SUBAPPLICATION GreenWhiteBackground2_AXC (* Hintergrundfarbe (TRUE -> Grün, FALSE -> Weiß) für 2 Objekte (AX-Adapter) (Kompakt) *)
  (* Standard: 61499-2 *)
  (* Version 1.0, 2026-07-21, franz, Meisterschulen am Ostbahnhof *)
  PACKAGE MyLib::sys;
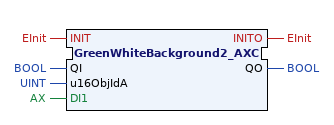
  EVENT_INPUT
    INIT : EInit; (* Initialization Request *)
  END_EVENT
  EVENT_OUTPUT
    INITO : EInit; (* Initialization Confirm *)
  END_EVENT
  VAR_INPUT
    QI : BOOL := TRUE; (* Quality Input - TRUE to enable service *)
    u16ObjIdA : UINT;
  END_VAR
  VAR_OUTPUT
    QO : BOOL; (* Quality Output - TRUE if service executed successfully *)
  END_VAR
  SOCKETS
    DI1 : adapter::types::unidirectional::AX;
  END_SOCKETS
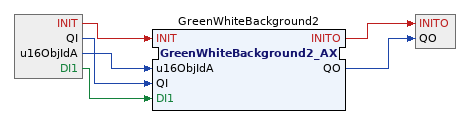
  SUBAPPS
    GreenWhiteBackground2 : MyLib::sys::GreenWhiteBackground2_AX;
  END_SUBAPPS
  EVENT_CONNECTIONS
    INIT TO GreenWhiteBackground2.INIT;
    GreenWhiteBackground2.INITO TO INITO;
  END_CONNECTIONS
  DATA_CONNECTIONS
    u16ObjIdA TO GreenWhiteBackground2.u16ObjIdA;
    QI TO GreenWhiteBackground2.QI;
    GreenWhiteBackground2.QO TO QO;
  END_CONNECTIONS
  ADAPTER_CONNECTIONS
    DI1 TO GreenWhiteBackground2.DI1;
  END_CONNECTIONS
END_SUBAPPLICATION
